// TIA Portal project "Proyecto_Marcha_Parada_20260708" (V13)

(* hardware
DEVICE "S7-1200 station_1"  S7-1200 Station
   slot 0: "Rack_0"  Rack  V1.0
   slot 1: "PLC_1"  CPU 1214C AC/DC/Rly  6ES7 214-1BE30-0XB0  V2.2
*)

// ===== PLC "PLC_1"  CPU 1214C AC/DC/Rly =====

VAR_GLOBAL   // PLC tag table "Tabla de variables estándar"
   "MARCHA" AT %I0.0 : Bool;
   "PARADA" AT %I0.1 : Bool;
   "MOTOR" AT %Q0.0 : Bool;
   "LUZ_PARADA" AT %Q0.1 : Bool;
   "LUZ_MARCHA" AT %Q0.2 : Bool;
END_VAR

ORGANIZATION_BLOCK "Main"   // OB1, LAD, ProgramCycle
TITLE = "Main Program Sweep (Cycle)"
{ S7_Optimized_Access := 'FALSE' }
VERSION : 0.1
BEGIN

REGION Network 1
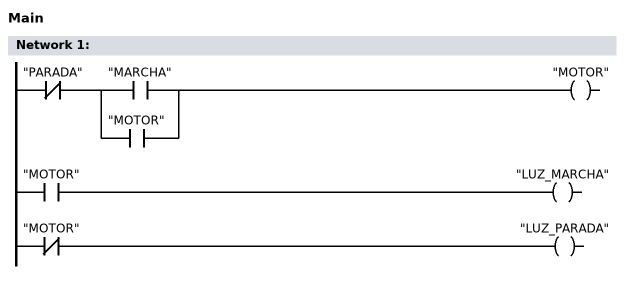
   RUNG wire#powerrail
      I_Contact( "PARADA" )
      wire#w1
      Contact( "MARCHA" )
      wire#w2
      Coil( "MOTOR" )
   END_RUNG
   RUNG wire#w1
      Contact( "MOTOR" )
   END_RUNG wire#w2
   RUNG wire#powerrail
      Contact( "MOTOR" )
      Coil( "LUZ_MARCHA" )
   END_RUNG
   RUNG wire#powerrail
      I_Contact( "MOTOR" )
      Coil( "LUZ_PARADA" )
   END_RUNG
   // the same network as SCL:
   "MOTOR" := NOT "PARADA" AND ("MARCHA" OR "MOTOR");
   "LUZ_MARCHA" := "MOTOR";
   "LUZ_PARADA" := NOT "MOTOR";
END_REGION
END_ORGANIZATION_BLOCK